// TIA Portal V20 export
Screen "190RobotCollision"  1276x673
  ScreenItem "矩形_6" at -3,69 size 1274x597  Type=HmiRectangle
  ScreenItem "Graphic view_13" at 324,87 size 634x531  Type=HmiGraphicView
  ScreenItem "Graphic view_5" at 101,0 size 472x35  Type=HmiGraphicView
  ScreenItem "Graphic view_9" at 0,7 size 472x35  Type=HmiGraphicView
  ScreenItem "Title_ScreenOverview_X390_Y2" at 438,5 size 551x57  Type=HmiTextBox
  ScreenItem "Line_Header_X0_Y64" at 0,64 size 1274x1  Type=HmiLine
  ScreenItem "permanentareaborderrectangle" at 0,0 size 0x0  Type=HmiRectangle
  ScreenItem "Button_Back" at 2,2 size 90x60  Type=HmiButton
  ScreenItem "Text_3" at 694,69 size 84x39  Type=HmiText
  ScreenItem "Text_4" at 627,514 size 84x39  Type=HmiText
  ScreenItem "Text_5" at 459,491 size 84x39  Type=HmiText
  ScreenItem "Text_6" at 476,68 size 84x39  Type=HmiText
  ScreenItem "Text_18" at 542,488 size 84x76  Type=HmiText
  ScreenItem "Graphic view_6" at 746,-206 size 60x30  Type=HmiGraphicView
  ScreenItem "Graphic view_7" at 746,-594 size 60x30  Type=HmiGraphicView
  ScreenItem "Graphic view_8" at 746,-982 size 60x30  Type=HmiGraphicView
  ScreenItem "Rectangle_5" at 893,75 size 164x112  Type=HmiRectangle
  ScreenItem "Text_71" at 885,70 size 174x35  Type=HmiText
  ScreenItem "Text_72" at 916,96 size 123x35  Type=HmiText
  ScreenItem "Text_73" at 930,124 size 88x35  Type=HmiText
  ScreenItem "Text_74" at 922,152 size 136x35  Type=HmiText
  ScreenItem "矩形_44" at 906,159 size 17x17  Type=HmiRectangle
  ScreenItem "矩形_45" at 906,132 size 17x17  Type=HmiRectangle
  ScreenItem "矩形_46" at 906,105 size 17x17  Type=HmiRectangle
  ScreenItem "Rectangle_6" at 809,415 size 164x222  Type=HmiRectangle
  ScreenItem "Text_75" at 801,410 size 174x35  Type=HmiText
  ScreenItem "Text_76" at 832,436 size 123x35  Type=HmiText
  ScreenItem "Text_77" at 846,464 size 88x35  Type=HmiText
  ScreenItem "Text_78" at 838,492 size 136x35  Type=HmiText
  ScreenItem "矩形_47" at 822,499 size 17x17  Type=HmiRectangle
  ScreenItem "矩形_48" at 822,472 size 17x17  Type=HmiRectangle
  ScreenItem "矩形_49" at 822,445 size 17x17  Type=HmiRectangle
  ScreenItem "Text_83" at 832,546 size 123x35  Type=HmiText
  ScreenItem "Text_84" at 801,520 size 174x35  Type=HmiText
  ScreenItem "矩形_53" at 822,555 size 17x17  Type=HmiRectangle
  ScreenItem "矩形_54" at 822,582 size 17x17  Type=HmiRectangle
  ScreenItem "矩形_55" at 822,609 size 17x17  Type=HmiRectangle
  ScreenItem "Text_85" at 838,602 size 136x35  Type=HmiText
  ScreenItem "Text_86" at 846,574 size 88x35  Type=HmiText
  ScreenItem "Graphic view_2" at 565,493 size 60x28  Type=HmiGraphicView
  ScreenItem "Graphic view_4" at 565,457 size 60x33  Type=HmiGraphicView
  ScreenItem "Text_1" at 562,409 size 84x73  Type=HmiText
  ScreenItem "Graphic view_11" at 88,0 size 410x35  Type=HmiGraphicView
  ScreenItem "Graphic view_12" at 0,7 size 410x35  Type=HmiGraphicView
  ScreenItem "Text_2" at 414,147 size 84x73  Type=HmiText
  ScreenItem "Text_9" at 414,378 size 84x73  Type=HmiText
  ScreenItem "Text_8" at 398,497 size 84x73  Type=HmiText
  ScreenItem "Rectangle_2" at 176,86 size 164x227  Type=HmiRectangle
  ScreenItem "Text_19" at 168,81 size 174x35  Type=HmiText
  ScreenItem "Text_20" at 199,107 size 123x35  Type=HmiText
  ScreenItem "Text_21" at 213,135 size 88x35  Type=HmiText
  ScreenItem "Text_22" at 205,163 size 136x35  Type=HmiText
  ScreenItem "矩形_8" at 189,170 size 17x17  Type=HmiRectangle
  ScreenItem "矩形_9" at 189,143 size 17x17  Type=HmiRectangle
  ScreenItem "矩形_10" at 189,116 size 17x17  Type=HmiRectangle
  ScreenItem "Graphic view_1" at 101,0 size 472x35  Type=HmiGraphicView
  ScreenItem "Graphic view_3" at 0,7 size 472x35  Type=HmiGraphicView
  ScreenItem "Text_23" at 414,90 size 84x73  Type=HmiText
  ScreenItem "Text_24" at 573,357 size 84x73  Type=HmiText
  ScreenItem "Text_25" at 759,86 size 84x73  Type=HmiText
  ScreenItem "Text_26" at 573,86 size 84x73  Type=HmiText
  ScreenItem "Graphic view_10" at 53,0 size 247x25  Type=HmiGraphicView
  ScreenItem "Graphic view_14" at 0,5 size 247x25  Type=HmiGraphicView
  ScreenItem "Text_27" at 375,606 size 84x39  Type=HmiText
  ScreenItem "Text_28" at 459,570 size 84x73  Type=HmiText
  ScreenItem "Rectangle_3" at 972,415 size 164x112  Type=HmiRectangle
  ScreenItem "Text_29" at 964,410 size 174x35  Type=HmiText
  ScreenItem "Text_30" at 995,436 size 123x35  Type=HmiText
  ScreenItem "Text_31" at 1009,464 size 88x35  Type=HmiText
  ScreenItem "Text_32" at 1001,492 size 136x35  Type=HmiText
  ScreenItem "矩形_11" at 985,499 size 17x17  Type=HmiRectangle
  ScreenItem "矩形_12" at 985,472 size 17x17  Type=HmiRectangle
  ScreenItem "矩形_13" at 985,445 size 17x17  Type=HmiRectangle
  ScreenItem "Text_7" at 165,192 size 174x35  Type=HmiText
  ScreenItem "Text_33" at 196,218 size 123x35  Type=HmiText
  ScreenItem "Text_34" at 210,246 size 88x35  Type=HmiText
  ScreenItem "Text_35" at 202,274 size 136x35  Type=HmiText
  ScreenItem "矩形_14" at 186,281 size 17x17  Type=HmiRectangle
  ScreenItem "矩形_15" at 186,254 size 17x17  Type=HmiRectangle
  ScreenItem "矩形_16" at 186,227 size 17x17  Type=HmiRectangle
  ScreenItem "Rectangle_1" at 219,394 size 164x224  Type=HmiRectangle
  ScreenItem "Text_10" at 211,389 size 174x35  Type=HmiText
  ScreenItem "Text_11" at 242,415 size 123x35  Type=HmiText
  ScreenItem "Text_12" at 256,443 size 88x35  Type=HmiText
  ScreenItem "Text_13" at 248,471 size 136x35  Type=HmiText
  ScreenItem "矩形_1" at 232,478 size 17x17  Type=HmiRectangle
  ScreenItem "矩形_2" at 232,451 size 17x17  Type=HmiRectangle
  ScreenItem "矩形_3" at 232,424 size 17x17  Type=HmiRectangle
  ScreenItem "Rectangle_4" at -427,725 size 164x112  Type=HmiRectangle
  ScreenItem "Text_14" at -435,720 size 174x35  Type=HmiText
  ScreenItem "Text_15" at -404,746 size 123x35  Type=HmiText
  ScreenItem "Text_16" at -390,774 size 88x35  Type=HmiText
  ScreenItem "Text_17" at -398,802 size 136x35  Type=HmiText
  ScreenItem "矩形_4" at -414,809 size 17x17  Type=HmiRectangle
  ScreenItem "矩形_5" at -414,782 size 17x17  Type=HmiRectangle
  ScreenItem "矩形_7" at -414,755 size 17x17  Type=HmiRectangle
  ScreenItem "Rectangle_7" at -1087,1044 size 164x112  Type=HmiRectangle
  ScreenItem "Text_36" at -1095,1039 size 174x35  Type=HmiText
  ScreenItem "Text_37" at -1064,1065 size 123x35  Type=HmiText
  ScreenItem "Text_38" at -1050,1093 size 88x35  Type=HmiText
  ScreenItem "Text_39" at -1058,1121 size 136x35  Type=HmiText
  ScreenItem "矩形_17" at -1074,1128 size 17x17  Type=HmiRectangle
  ScreenItem "矩形_18" at -1074,1101 size 17x17  Type=HmiRectangle
  ScreenItem "矩形_19" at -1074,1074 size 17x17  Type=HmiRectangle
  ScreenItem "Rectangle_8" at -1747,1363 size 164x112  Type=HmiRectangle
  ScreenItem "Text_40" at -1724,1384 size 123x35  Type=HmiText
  ScreenItem "Text_41" at -1710,1412 size 88x35  Type=HmiText
  ScreenItem "Text_42" at -1718,1440 size 136x35  Type=HmiText
  ScreenItem "矩形_20" at -1734,1447 size 17x17  Type=HmiRectangle
  ScreenItem "矩形_21" at -1734,1420 size 17x17  Type=HmiRectangle
  ScreenItem "矩形_22" at -1734,1393 size 17x17  Type=HmiRectangle
  ScreenItem "Rectangle_9" at -2407,1682 size 164x112  Type=HmiRectangle
  ScreenItem "Text_43" at -2415,1677 size 174x35  Type=HmiText
  ScreenItem "Text_44" at -2384,1703 size 123x35  Type=HmiText
  ScreenItem "Text_45" at -2370,1731 size 88x35  Type=HmiText
  ScreenItem "Text_46" at -2378,1759 size 136x35  Type=HmiText
  ScreenItem "矩形_23" at -2394,1766 size 17x17  Type=HmiRectangle
  ScreenItem "矩形_24" at -2394,1739 size 17x17  Type=HmiRectangle
  ScreenItem "矩形_25" at -2394,1712 size 17x17  Type=HmiRectangle
  ScreenItem "Rectangle_10" at 595,548 size 164x112  Type=HmiRectangle
  ScreenItem "Text_47" at 587,543 size 174x35  Type=HmiText
  ScreenItem "Text_48" at 618,569 size 123x35  Type=HmiText
  ScreenItem "Text_49" at 632,597 size 88x35  Type=HmiText
  ScreenItem "Text_50" at 624,625 size 136x35  Type=HmiText
  ScreenItem "矩形_26" at 608,632 size 17x17  Type=HmiRectangle
  ScreenItem "矩形_27" at 608,605 size 17x17  Type=HmiRectangle
  ScreenItem "矩形_28" at 608,578 size 17x17  Type=HmiRectangle
  ScreenItem "Text_51" at 215,499 size 174x35  Type=HmiText
  ScreenItem "Text_52" at 246,525 size 123x35  Type=HmiText
  ScreenItem "Text_53" at 260,553 size 88x35  Type=HmiText
  ScreenItem "Text_54" at 252,581 size 136x35  Type=HmiText
  ScreenItem "矩形_29" at 236,588 size 17x17  Type=HmiRectangle
  ScreenItem "矩形_30" at 236,561 size 17x17  Type=HmiRectangle
  ScreenItem "矩形_31" at 236,534 size 17x17  Type=HmiRectangle
